// TIA Portal V21 export
// export: Created 2026-11-10T19:11:38.3560932Z, ExportSetting WithDefaults, DisplayName Totally Integrated Automation Portal, DisplayVersion V21 Update 3, DisplayName STEP 7 Professional, DisplayVersion V21 Update 3, DisplayName STEP 7 Safety, DisplayVersion V21, DisplayName Tech WebApplication, DisplayVersion V21, DisplayName WinCC Basic/Comfort/Advanced, DisplayVersion V21 Update 3, DisplayName WinCC Unified, DisplayVersion V21 Update 3
DATA_BLOCK "DB_SMC"   // DB26
// stored: AutoNumber true, DBAccessibleFromOPCUA true, DBAccessibleFromWebserver true, InstanceOfName SMC, OfSystemLibElement SMC, OfSystemLibVersion 2.1
"SMC"
   // VAR_INPUT
   //    IN_BIT0 : Bool;
   //    IN_BIT1 : Bool;
   //    IN_BIT2 : Bool;
   //    IN_BIT3 : Bool;
   //    IN_BIT4 : Bool;
   //    IN_BIT5 : Bool;
   //    IN_BIT6 : Bool;
   //    IN_BIT7 : Bool;
   //    IN_BIT8 : Bool;
   //    IN_BIT9 : Bool;
   //    IN_BIT10 : Bool;
   //    IN_BIT11 : Bool;
   //    IN_BIT12 : Bool;
   //    IN_BIT13 : Bool;
   //    IN_BIT14 : Bool;
   //    IN_BIT15 : Bool;
   // END_VAR
   // VAR_OUTPUT
   //    OUT : Bool;
   //    ERR_CODE : Word;
   //    OUT_STEP : Byte;
   // END_VAR
   // VAR
   //    LAST : Byte;
   //    CMP_VAL : Array[0..15, 0..15] of Bool;
   // END_VAR
BEGIN
END_DATA_BLOCK
